{attribute 'qualified_only'}
// Robot CM sizing (Annex I). The user channel is a small DECLARED set, not a
// mailbox: eight signals cover a gripper, a program flag or two and a counter,
// and a bound is what keeps it from becoming a second command surface.
VAR_GLOBAL CONSTANT
    MAX_USER_SIGNALS : INT := 8;
    MAX_JOG_AXES     : INT := 7;   // joint jog addresses axes 1..7; Cartesian/tool 1..6
    // Declared one-press manual moves (M_DeclareManualMove). Eight, because the
    // catalog holds MAX_CMD_CATALOG (12) and the type publishes four of its own:
    // two held jogs, the brake test and the safe reference run.
    MAX_MANUAL_MOVES : INT := 8;
    // Catalog value of manual move n is MANUAL_MOVE_BASE + n: clear of every
    // E_RobotCommand value, so a press can never be read as another command.
    MANUAL_MOVE_BASE : DINT := 100;
END_VAR

(* stored: Version 1.1.0.1, ProductVersion 3.1.4024.12
   GVL PL_Robot: Id {60011b9f-d90e-42a5-b6b6-823816846d87} *)
